// TIA Portal V20 export
ORGANIZATION_BLOCK "T2_Ciclo_Nuevos"   // OB126, LAD, ProgramCycle
TITLE = T2_Ciclo_Nuevos
{ S7_Optimized_Access := 'TRUE' }
AUTHOR : IA
FAMILY : PRUEBA
VERSION : 0.1
// Prueba IA 3: una FC por construcción nueva
// stored: AutoNumber false, IsIECCheckEnabled false, SetENOAutomatically false
   VAR_INPUT
      Initial_Call : Bool;
      Remanence : Bool;
   END_VAR
BEGIN

REGION Network 1: Contador de vida
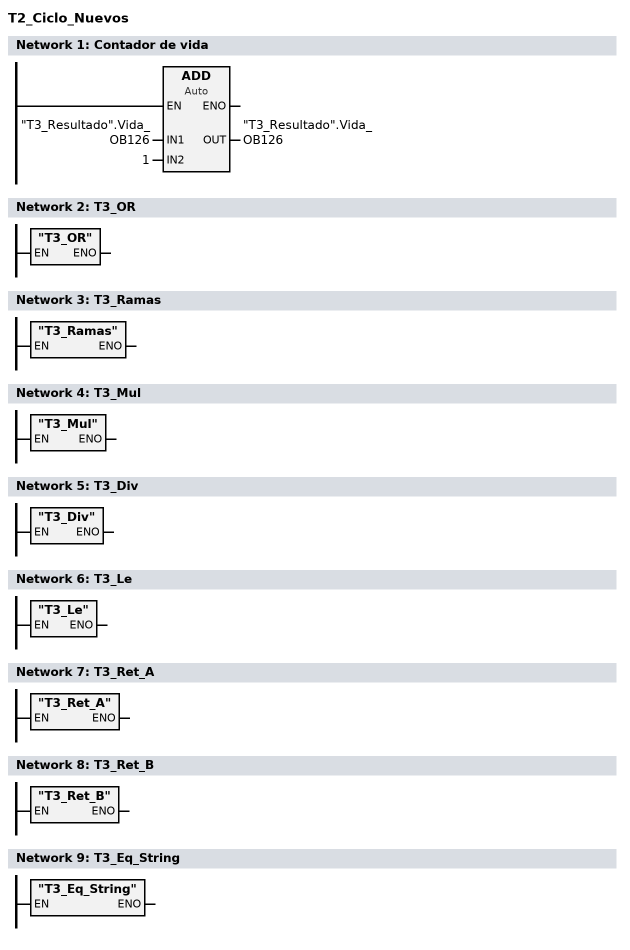
   RUNG wire#powerrail
      Add(in1 := "T3_Resultado".Vida_OB126, in2 := 1, out => "T3_Resultado".Vida_OB126)
   END_RUNG
   // the same network as SCL:
   "T3_Resultado".Vida_OB126 := "T3_Resultado".Vida_OB126 + 1;
END_REGION

REGION Network 2: T3_OR
   RUNG wire#powerrail
      "T3_OR"()
   END_RUNG
   // the same network as SCL:
   "T3_OR"();
END_REGION

REGION Network 3: T3_Ramas
   RUNG wire#powerrail
      "T3_Ramas"()
   END_RUNG
   // the same network as SCL:
   "T3_Ramas"();
END_REGION

REGION Network 4: T3_Mul
   RUNG wire#powerrail
      "T3_Mul"()
   END_RUNG
   // the same network as SCL:
   "T3_Mul"();
END_REGION

REGION Network 5: T3_Div
   RUNG wire#powerrail
      "T3_Div"()
   END_RUNG
   // the same network as SCL:
   "T3_Div"();
END_REGION

REGION Network 6: T3_Le
   RUNG wire#powerrail
      "T3_Le"()
   END_RUNG
   // the same network as SCL:
   "T3_Le"();
END_REGION

REGION Network 7: T3_Ret_A
   RUNG wire#powerrail
      "T3_Ret_A"()
   END_RUNG
   // the same network as SCL:
   "T3_Ret_A"();
END_REGION

REGION Network 8: T3_Ret_B
   RUNG wire#powerrail
      "T3_Ret_B"()
   END_RUNG
   // the same network as SCL:
   "T3_Ret_B"();
END_REGION

REGION Network 9: T3_Eq_String
   RUNG wire#powerrail
      "T3_Eq_String"()
   END_RUNG
   // the same network as SCL:
   "T3_Eq_String"();
END_REGION
END_ORGANIZATION_BLOCK
